(* IEC 61131-3 sources: bcs-engineering-dsl/language/test/generating/enum_test/expected, 3 files *)

(* ---- Mode.st ---- *)
{attribute 'qualified_only'}
{attribute 'strict'}
TYPE Mode :
(
    OFF := 0,
    ECO := 1,
    COMFORT := 2
);
END_TYPE

(* ---- MAIN_decl.st ---- *)
PROGRAM MAIN
VAR
    windowContact_value AT %I*: BOOL; (* Input channel from hardware *)
    previousMode: Mode := Mode.OFF;
    TestUnit_currentMode: Mode := Mode.OFF;
END_VAR

(* ---- MAIN_impl.st ---- *)
// Control Unit 'TestUnit'
IF TestUnit_currentMode = Mode.ECO THEN
    previousMode := TestUnit_currentMode;
    TestUnit_currentMode := Mode.COMFORT;
END_IF;
